INTERFACE I_Axis

METHOD Enable : E_PROGRESS
VAR_INPUT
END_VAR
END_METHOD

METHOD Disable : E_PROGRESS
VAR_INPUT
END_VAR
END_METHOD

METHOD Reset : E_PROGRESS
VAR_INPUT
END_VAR
END_METHOD

METHOD Home : E_PROGRESS
VAR_INPUT
END_VAR
END_METHOD

METHOD MoveAbsolute : E_PROGRESS
VAR_INPUT
    lrPosition : LREAL;   // [units]
    lrVelocity : LREAL;   // [units/s]
END_VAR
END_METHOD

METHOD MoveRelative : E_PROGRESS
VAR_INPUT
    lrDistance : LREAL;   // [units]
    lrVelocity : LREAL;   // [units/s]
END_VAR
END_METHOD

METHOD MoveVelocity : E_PROGRESS
VAR_INPUT
    lrVelocity : LREAL;   // [units/s] signed
END_VAR
END_METHOD

METHOD Jog : E_PROGRESS
VAR_INPUT
    xForward   : BOOL;
    xReverse   : BOOL;
    lrVelocity : LREAL;   // magnitude [units/s]
END_VAR
END_METHOD

METHOD MoveFollow : E_PROGRESS
VAR_INPUT
    lrPosition : LREAL;   // [units] - online re-targetable
    lrVelocity : LREAL;   // [units/s]
END_VAR
END_METHOD

METHOD Stop : E_PROGRESS
VAR_INPUT
END_VAR
END_METHOD

PROPERTY Position : LREAL
GET
END_GET
END_PROPERTY

PROPERTY Enabled : BOOL
GET
END_GET
END_PROPERTY

END_INTERFACE

(* stored: Version 1.1.0.1
   Itf I_Axis: Id {9993b2d1-1971-5037-9cc4-3616bff67ba3}
   Method Enable: Id {a91b16c2-4aac-55a7-8408-a1d51b752d8e}
   Method Disable: Id {ff6e472e-7452-5f39-8d7c-a260cab339ff}
   Method Reset: Id {c71cdb91-579b-5a8c-9f54-6d76c0afa2b4}
   Method Home: Id {fe930bd5-867a-551e-9e84-f3c4c864c429}
   Method MoveAbsolute: Id {3ddce93d-0461-53af-a1ea-091e13ee7098}
   Method MoveRelative: Id {6d8a97c0-823b-5bd6-bc3a-36688fc5a9da}
   Method MoveVelocity: Id {569f99f6-0a71-5e1d-9355-5a679ae6d8ed}
   Method Jog: Id {5c5a5a2a-9cec-5c0a-b230-b1d24afc8046}
   Method MoveFollow: Id {d314823a-64ff-57ef-90fe-f60b1d7a1d6a}
   Method Stop: Id {1b6ffba0-5b04-5df9-ac0c-b45290944e69}
   Property Position: Id {53cb5025-8f91-575a-9ec0-7a93eb759990}
   Get Get: Id {e136aa8c-8ca8-55c9-8d8c-145384a8e27f}
   Property Enabled: Id {41b72ac1-7553-5dc7-ab72-f15a4e10e403}
   Get Get: Id {fd6d7d5e-8a8d-5534-8a63-9d56a3d4bc1f} *)
